(* IEC 61131-3 sources: ICSPrism/benchmarks, 8 files *)

(* ---- harness_test.st ---- *)
FUNCTION_BLOCK Counter
VAR_INPUT
    Increment : INT;
    Reset     : BOOL;
END_VAR
VAR
    Value     : INT;
    TotalCalls: INT;
END_VAR

TotalCalls := TotalCalls + 1;
IF Reset THEN
    Value := 0;
ELSE
    Value := Value + Increment;
END_IF
END_FUNCTION_BLOCK

PROGRAM HarnessTest
VAR_INPUT
    A        : INT;       (* i16 scalar input           *)
    B        : INT;       (* i16 scalar input           *)
    Flag     : BOOL;      (* i8  boolean input          *)
    Index    : INT;       (* i16 used as array index    *)
END_VAR
VAR
    Sum      : INT;       (* A + B each cycle           *)
    Product  : DINT;      (* A * B, wider type          *)
    Buf      : ARRAY[0..15] OF INT;  (* 16-element buffer *)
    C        : Counter;   (* nested function block      *)
    CycleNum : INT;       (* increments every scan      *)
END_VAR

(* Simple deterministic behavior easy to verify *)
CycleNum := CycleNum + 1;
Sum      := A + B;
Product  := A * B;

(* Bounded array write — safe when 0 <= Index <= 15 *)
IF Index >= 0 AND Index <= 15 THEN
    Buf[Index] := Sum;
END_IF

(* Drive the nested counter *)
C(Increment := A, Reset := Flag);

END_PROGRAM

(* ---- harness_test_buggy.st ---- *)
FUNCTION_BLOCK Counter
VAR_INPUT
    Increment : INT;
    Reset     : BOOL;
END_VAR
VAR
    Value     : INT;
    TotalCalls: INT;
END_VAR

TotalCalls := TotalCalls + 1;
IF Reset THEN
    Value := 0;
ELSE
    Value := Value + Increment;
END_IF
END_FUNCTION_BLOCK

PROGRAM HarnessTest
VAR_INPUT
    A        : INT;       (* i16 scalar input           *)
    B        : INT;       (* i16 scalar input           *)
    Flag     : BOOL;      (* i8  boolean input          *)
    Index    : INT;       (* i16 used as array index    *)
END_VAR
VAR
    Sum      : INT;       (* A + B each cycle           *)
    Product  : DINT;      (* A * B, wider type          *)
    Buf      : ARRAY[0..15] OF INT;  (* 16-element buffer *)
    C        : Counter;   (* nested function block      *)
    CycleNum : INT;       (* increments every scan      *)
END_VAR

(* Simple deterministic behavior easy to verify *)
CycleNum := CycleNum + 1;
Sum      := A + B;
Product  := A * B;

(* Bounded array write — safe when 0 <= Index <= 15 *)
IF Index >= 0 OR Index <= 15 THEN
    Buf[Index] := Sum;
END_IF

(* Drive the nested counter *)
C(Increment := A, Reset := Flag);

END_PROGRAM

(* ---- pipeline_controller.st ---- *)
{external}
FUNCTION prism_bug_abort_if : DINT
VAR_INPUT
    should_abort : DINT;
    bug_id       : DINT;
END_VAR
END_FUNCTION

// pipeline_controller — industrial pipeline fill process controller
//
// Bug: Buffer[FillHead] OOB write when FillHead >= 64 (Buffer is [0..63]).
//
// Why this benchmark is decisively harder for input-only fuzzing:
//
//   (1) FillHead is NEVER compared against 64 — it appears only as an array
//       index. trace-cmp has zero visibility into its growth toward 64.
//
//   (2) TWO-DIMENSIONAL ZONE DECAY with 8 zones:
//       FillHead [0,63] is split into 8 zones of 8. Each zone simultaneously
//       requires (PumpRate + ValvePos) AND PipeTemp to be in specific windows.
//       The windows are arranged so that NO fixed (PumpRate, ValvePos, PipeTemp)
//       triple satisfies all 8 zones — and several consecutive zone transitions
//       require coordinated simultaneous changes in multiple inputs.
//
//       Zone 0 [FH  0- 7]: PVsum [60,90]   PipeTemp [50,65]
//       Zone 1 [FH  8-15]: PVsum [80,110]  PipeTemp [62,77]   PVsum up, temp up
//       Zone 2 [FH 16-23]: PVsum [70,100]  PipeTemp [72,87]   PVsum back, temp up
//       Zone 3 [FH 24-31]: PVsum [55, 85]  PipeTemp [65,80]   PVsum down, temp down
//       Zone 4 [FH 32-39]: PVsum [95,125]  PipeTemp [55,70]   PVsum jumps (gap!)
//       Zone 5 [FH 40-47]: PVsum [65, 95]  PipeTemp [78,93]   PVsum down, temp jumps (gap!)
//       Zone 6 [FH 48-55]: PVsum [85,115]  PipeTemp [52,67]   PVsum up, temp folds back (gap!)
//       Zone 7 [FH 56-63]: PVsum [75,105]  PipeTemp [63,78]   PVsum down, temp up
//
//       Critical transitions with NO input overlap between zones:
//         3→4: PVsum must jump from ≤85 to ≥95 (9-unit gap)
//         4→5: PipeTemp must jump from ≤70 to ≥78 while PVsum drops
//         5→6: PipeTemp must drop from ≥78 to ≤67 (fold-back of ~20 units)
//
//   (3) 7 inputs (vs 4 in valve_sequencer) give the custom mutator a richer
//       space: for each zone, PumpRate AND ValvePos AND PipeTemp must be set
//       correctly — three bytes to coordinate, not one.
//
//   (4) Decay is -6 per bad cycle vs +1 advance per 4th qualifying cycle.
//       Random inputs decay FillHead rapidly; only sustained zone-correct
//       inputs allow growth. Without FillHead state signal, the fuzzer cannot
//       know which zone it is in or which transition is approaching.
//
//   (5) Two pre-fill phases (PRIME, FLOW) are guided by trace-cmp and add
//       ~80 cycles of required navigation before FILL begins.
//
// Phase path:
//   IDLE  → Cmd = 1
//   PRIME → PrimeScore >= 8   (every 3rd phase-cycle, combined sum, decay-2) ~30+ cycles
//   FLOW  → FluxScore >= 8    (combined PipeTemp+CoolantRate, halved/11cy)   ~50+ cycles
//   FILL  → FillHead reaches 64 (every 4th qualifying cycle, 8-zone 2D decay) ~300+ cycles
//
// Key variables for state signal: Phase, PrimeScore, FluxScore,
//   FlowAccum, PressAccum, TempAccum, FillHead.
// FillHead is the only one invisible to trace-cmp.
// (PVsum = PumpRate + ValvePos) zone requirements make the state signal
// especially valuable: the fuzzer must know FillHead to know which inputs
// to set, which trace-cmp cannot determine from TempIn comparisons alone.

VAR_GLOBAL CONSTANT
    PHASE_IDLE  : SINT := 0;
    PHASE_PRIME : SINT := 1;
    PHASE_FLOW  : SINT := 2;
    PHASE_FILL  : SINT := 3;
END_VAR

PROGRAM PLC_PRG
VAR_INPUT
    PumpRate    : INT  := 0;
    ValvePos    : INT  := 0;
    PipeTemp    : INT  := 0;
    BackPressure: INT  := 0;
    FeedConc    : INT  := 0;
    CoolantRate : INT  := 0;
    Cmd         : SINT := 0;
END_VAR
VAR
    Ctrl : PipelineCtrl;
END_VAR

Ctrl(
    PumpRate     := PumpRate,
    ValvePos     := ValvePos,
    PipeTemp     := PipeTemp,
    BackPressure := BackPressure,
    FeedConc     := FeedConc,
    CoolantRate  := CoolantRate,
    Cmd          := Cmd
);

END_PROGRAM

FUNCTION_BLOCK PipelineCtrl
VAR_INPUT
    PumpRate    : INT;
    ValvePos    : INT;
    PipeTemp    : INT;
    BackPressure: INT;
    FeedConc    : INT;
    CoolantRate : INT;
    Cmd         : SINT;
END_VAR
VAR_OUTPUT
    Status      : SINT;
END_VAR
VAR
    Phase        : SINT := PHASE_IDLE;
    CycleCount   : INT  := 0;
    // PRIME phase
    PrimeCycles  : INT  := 0;
    PrimeScore   : INT  := 0;
    // FLOW phase
    FluxScore    : INT  := 0;
    FluxSum      : INT  := 0;
    // FILL phase accumulators
    FlowAccum    : INT  := 0;
    PressAccum   : INT  := 0;
    TempAccum    : INT  := 0;
    PhaseCounter : INT  := 0;
    // Hidden OOB counter — NEVER compared against 64, only used as array index
    FillHead     : INT  := 0;
    // OOB write target
    Buffer       : ARRAY[0..63] OF INT;
    PVsum        : INT  := 0;
    i            : INT;
END_VAR

CycleCount := CycleCount + 1;

CASE Phase OF

    PHASE_IDLE:
        IF Cmd = 1 THEN
            FOR i := 0 TO 63 DO
                Buffer[i] := 0;
            END_FOR;
            PrimeCycles  := 0;
            PrimeScore   := 0;
            FluxScore    := 0;
            FlowAccum    := 0;
            PressAccum   := 0;
            TempAccum    := 0;
            PhaseCounter := 0;
            FillHead     := 0;
            PVsum        := 0;
            Phase        := PHASE_PRIME;
        END_IF;

    PHASE_PRIME:
        // Combined PumpRate+BackPressure sum forces simultaneous tuning of
        // two inputs. trace-cmp sees the sum, not individual contributions.
        // Only every 3rd phase-cycle counts; decay-2 forces sustained inputs.
        PrimeCycles := PrimeCycles + 1;
        PVsum := PumpRate + BackPressure;

        IF PrimeCycles MOD 3 = 0 THEN
            IF PVsum >= 80 AND PVsum <= 160 AND ValvePos >= 15 AND ValvePos <= 60 THEN
                PrimeScore := PrimeScore + 1;
            ELSE
                IF PrimeScore > 1 THEN
                    PrimeScore := PrimeScore - 2;
                ELSE
                    PrimeScore := 0;
                END_IF;
            END_IF;
        END_IF;

        IF PrimeScore >= 8 THEN
            Phase := PHASE_FLOW;
        END_IF;

    PHASE_FLOW:
        // Combined PipeTemp + CoolantRate sum partially hides which input is
        // responsible. Halved every 11 global cycles — forces sustained inputs.
        FluxSum := PipeTemp + CoolantRate;

        IF FluxSum >= 80 AND FluxSum <= 160 AND FeedConc >= 20 AND FeedConc <= 70 THEN
            FluxScore := FluxScore + 1;
        ELSE
            IF FluxScore > 1 THEN
                FluxScore := FluxScore - 2;
            ELSE
                FluxScore := 0;
            END_IF;
        END_IF;

        IF CycleCount MOD 11 = 0 AND FluxScore > 0 THEN
            FluxScore := FluxScore / 2;
        END_IF;

        IF FluxScore >= 8 THEN
            Phase := PHASE_FILL;
        END_IF;

    PHASE_FILL:
        PhaseCounter := PhaseCounter + 1;

        // Three accumulator channels — all visible to trace-cmp, which guides
        // the fuzzer into FILL and maintains channel health.

        IF PumpRate >= 40 AND PumpRate <= 90 THEN
            FlowAccum := FlowAccum + 1;
        ELSE
            IF FlowAccum > 1 THEN
                FlowAccum := FlowAccum - 2;
            ELSE
                FlowAccum := 0;
            END_IF;
        END_IF;

        IF BackPressure >= 30 AND BackPressure <= 80 THEN
            PressAccum := PressAccum + 1;
        ELSE
            IF PressAccum > 0 THEN
                PressAccum := PressAccum - 1;
            END_IF;
        END_IF;

        // TempAccum window [50,100] — all zone PipeTemp windows are subsets
        // of this range, so zone requirements always keep TempAccum healthy.
        IF PipeTemp >= 50 AND PipeTemp <= 100 THEN
            TempAccum := TempAccum + 1;
        ELSE
            IF TempAccum > 1 THEN
                TempAccum := TempAccum - 2;
            ELSE
                TempAccum := 0;
            END_IF;
        END_IF;

        // FillHead advances every 4th qualifying cycle.
        // FillHead is NEVER compared against 64 — only appears as array index.
        IF FlowAccum > 6 AND PressAccum > 5 AND TempAccum > 6 THEN
            IF PhaseCounter MOD 4 = 0 THEN
                FillHead := FillHead + 1;
            END_IF;
        END_IF;

        // TWO-DIMENSIONAL ZONE DECAY — the decisive state-signal barrier:
        //
        // FillHead [0,63] is partitioned into 8 zones of 8. Each zone requires
        // BOTH (PumpRate + ValvePos) AND PipeTemp to be in specific windows.
        // These two conditions must be met simultaneously every cycle or FillHead
        // decays by 6 — erasing up to 6 accumulated advances in one bad cycle.
        //
        // Critical transitions (no overlap between adjacent zones):
        //   3→4: PVsum must jump from ≤85 to ≥95 — 9-unit gap, must coordinate
        //         PumpRate AND ValvePos inputs at exactly the right cycle
        //   4→5: PipeTemp must jump ≥8 units while PVsum drops ≥30 units
        //   5→6: PipeTemp must drop ≥11 units (fold-back)
        //
        // trace-cmp instruments PVsum and PipeTemp comparisons but the required
        // windows change with FillHead (state, not input). An input-only fuzzer
        // receives conflicting gradients: e.g., PVsum should be high for zone 4
        // but low for zones 0, 2, 3, 5. Only the key-state signal on FillHead
        // reveals which zone is currently active.
        //
        // A custom mutator with FillHead signal can look up the current zone and
        // set PumpRate, ValvePos, AND PipeTemp precisely — three bytes at once.
        PVsum := PumpRate + ValvePos;

        IF FillHead < 8 THEN
            // Zone 0: PVsum [60,90], PipeTemp [50,65]
            IF PVsum < 60 OR PVsum > 90 OR PipeTemp < 50 OR PipeTemp > 65 THEN
                IF FillHead > 5 THEN
                    FillHead := FillHead - 6;
                ELSE
                    FillHead := 0;
                END_IF;
            END_IF;
        ELSIF FillHead < 16 THEN
            // Zone 1: PVsum [80,110], PipeTemp [62,77]
            IF PVsum < 80 OR PVsum > 110 OR PipeTemp < 62 OR PipeTemp > 77 THEN
                IF FillHead > 5 THEN
                    FillHead := FillHead - 6;
                ELSE
                    FillHead := 0;
                END_IF;
            END_IF;
        ELSIF FillHead < 24 THEN
            // Zone 2: PVsum [70,100], PipeTemp [72,87]
            IF PVsum < 70 OR PVsum > 100 OR PipeTemp < 72 OR PipeTemp > 87 THEN
                IF FillHead > 5 THEN
                    FillHead := FillHead - 6;
                ELSE
                    FillHead := 0;
                END_IF;
            END_IF;
        ELSIF FillHead < 32 THEN
            // Zone 3: PVsum [55,85], PipeTemp [65,80]
            IF PVsum < 55 OR PVsum > 85 OR PipeTemp < 65 OR PipeTemp > 80 THEN
                IF FillHead > 5 THEN
                    FillHead := FillHead - 6;
                ELSE
                    FillHead := 0;
                END_IF;
            END_IF;
        ELSIF FillHead < 40 THEN
            // Zone 4: PVsum [95,125], PipeTemp [55,70]
            // *** GAP from zone 3: PVsum must jump from ≤85 to ≥95 ***
            IF PVsum < 95 OR PVsum > 125 OR PipeTemp < 55 OR PipeTemp > 70 THEN
                IF FillHead > 5 THEN
                    FillHead := FillHead - 6;
                ELSE
                    FillHead := 0;
                END_IF;
            END_IF;
        ELSIF FillHead < 48 THEN
            // Zone 5: PVsum [65,95], PipeTemp [78,93]
            // *** GAP from zone 4: PipeTemp must jump from ≤70 to ≥78 ***
            IF PVsum < 65 OR PVsum > 95 OR PipeTemp < 78 OR PipeTemp > 93 THEN
                IF FillHead > 5 THEN
                    FillHead := FillHead - 6;
                ELSE
                    FillHead := 0;
                END_IF;
            END_IF;
        ELSIF FillHead < 56 THEN
            // Zone 6: PVsum [85,115], PipeTemp [52,67]
            // *** GAP from zone 5: PipeTemp must drop from ≥78 to ≤67 ***
            IF PVsum < 85 OR PVsum > 115 OR PipeTemp < 52 OR PipeTemp > 67 THEN
                IF FillHead > 5 THEN
                    FillHead := FillHead - 6;
                ELSE
                    FillHead := 0;
                END_IF;
            END_IF;
        ELSE
            // Zone 7: PVsum [75,105], PipeTemp [63,78]
            IF PVsum < 75 OR PVsum > 105 OR PipeTemp < 63 OR PipeTemp > 78 THEN
                IF FillHead > 5 THEN
                    FillHead := FillHead - 6;
                ELSE
                    FillHead := 0;
                END_IF;
            END_IF;
        END_IF;

        // OOB write: Buffer is [0..63] (64 elements).
        // FillHead >= 64 writes out of bounds.
        // FillHead appears ONLY here — no comparison against 64 anywhere.
        Buffer[FillHead] := CycleCount;
        IF FillHead > 63 THEN
            prism_bug_abort_if(1, 9001);
        END_IF;

END_CASE;

Status := Phase;

END_FUNCTION_BLOCK

(* ---- pump_controller.st ---- *)
{external}
FUNCTION prism_bug_abort_if : DINT
VAR_INPUT
    should_abort : DINT;
    bug_id       : DINT;
END_VAR
END_FUNCTION

VAR_GLOBAL CONSTANT
    MODE_INIT  : SINT := 0;
    MODE_IDLE  : SINT := 1;
    MODE_ARMED : SINT := 2;
    MODE_RUN   : SINT := 3;
    MODE_FAULT : SINT := 4;
END_VAR

PROGRAM PLC_PRG
VAR_INPUT
    CmdArm    : BOOL := FALSE;
    CmdStart  : BOOL := FALSE;
    CmdReset  : BOOL := FALSE;
    Pressure  : INT := 0;
    Temp      : INT := 0;
END_VAR
VAR
    Controller : PumpController;
END_VAR

Controller(
    CmdArm := CmdArm,
    CmdStart := CmdStart,
    CmdReset := CmdReset,
    Pressure := Pressure,
    Temp := Temp
);

END_PROGRAM

FUNCTION_BLOCK PumpController
VAR_INPUT
    CmdArm    : BOOL;
    CmdStart  : BOOL;
    CmdReset  : BOOL;
    Pressure  : INT;
    Temp      : INT;
END_VAR
VAR
    Mode          : SINT := MODE_INIT;
    CycleCount    : INT := 0;
    PressureScore : INT := 0;
    ArmedCycles   : INT := 0;
    Offset        : INT := 0;
    Buffer        : ARRAY[0..7] OF INT;
    i             : INT;
END_VAR
VAR_OUTPUT
    Status        : SINT;
END_VAR

CycleCount := CycleCount + 1;

CASE Mode OF

    MODE_INIT:
        FOR i := 0 TO 7 DO
            Buffer[i] := 0;
        END_FOR;
        PressureScore := 0;
        ArmedCycles := 0;
        Offset := 0;
        Mode := MODE_IDLE;

    MODE_IDLE:
        IF CmdReset THEN
            PressureScore := 0;
            ArmedCycles := 0;
            Offset := 0;
        END_IF;

        IF CmdArm THEN
            Mode := MODE_ARMED;
            ArmedCycles := 0;
        END_IF;

    MODE_ARMED:
        ArmedCycles := ArmedCycles + 1;

        IF CmdReset THEN
            Mode := MODE_IDLE;
            PressureScore := 0;
            ArmedCycles := 0;
            Offset := 0;
        ELSIF CmdStart AND ArmedCycles >= 3 THEN
            Mode := MODE_RUN;
        END_IF;

    MODE_RUN:
        IF Pressure > 70 THEN
            PressureScore := PressureScore + 1;
        END_IF;

        IF Temp > 50 AND Temp < 60 THEN
            Offset := Offset + 1;
        END_IF;

        IF PressureScore >= 4 THEN
            Buffer[0] := Buffer[0] + 1;
        END_IF;

        IF Buffer[0] > 2 THEN
            Buffer[1] := Buffer[1] + 1;
        END_IF;

        // Deliberate deep bug:
        // Requires entering RUN, then building enough history so Offset becomes large.
        // Input-only fuzzing with frequent resets should struggle more than stateful fuzzing.
        IF Buffer[1] > 1 THEN
            Buffer[Offset] := 1234;
            IF Offset > 7 THEN
                prism_bug_abort_if(1, 9001);
            END_IF;
        END_IF;

        IF CmdReset THEN
            Mode := MODE_IDLE;
            PressureScore := 0;
            ArmedCycles := 0;
            Offset := 0;
        END_IF;

        IF Temp > 90 THEN
            Mode := MODE_FAULT;
        END_IF;

    MODE_FAULT:
        IF CmdReset THEN
            Mode := MODE_IDLE;
            PressureScore := 0;
            ArmedCycles := 0;
            Offset := 0;
        END_IF;

END_CASE;

Status := Mode;

END_FUNCTION_BLOCK

(* ---- scan_cycle_aircraft_oobr.st ---- *)
VAR_GLOBAL CONSTANT
    SS_INITIALIZE: SINT := 0;
    SS_STEP: SINT := 1;
    SS_FIN: SINT := 2;
END_VAR

PROGRAM PLC_PRG
VAR_INPUT
	In: ARRAY[0..7] OF LREAL := [3.0, 2.0, 3.0, 4.0, 1.0, 0.0, -1.0, 2.5];
    ssMethodType: SINT := SS_INITIALIZE;
END_VAR
VAR
	Out: ARRAY[0..1] OF LREAL;
    Code: Code;
END_VAR

// Harness simulation
Code(In, ssMethodType);

END_PROGRAM

FUNCTION_BLOCK Code
VAR_IN_OUT
    InRecv: ARRAY[0..7] OF LREAL;
    ssMethodType: SINT;
END_VAR
VAR
	offset: DWORD;
    CycleCount: INT;
	wGust: LREAL;
    qGust: LREAL;
    iter: INT;
	In: ARRAY[0..64] OF LREAL;
END_VAR
VAR_OUTPUT
    Out: ARRAY[0..1] OF LREAL;
END_VAR

// Complex branching logic
CASE ssMethodType OF

    SS_INITIALIZE:
        // Initialize memory
        FOR iter := 0 TO 64 DO
            In[iter] := 0.0;
        END_FOR;
        ssMethodType := SS_STEP;

    SS_STEP:

        // Copy Inputs
        CycleCount := CycleCount + 1;
        MemCpy(ADR(In), ADR(InRecv), offset);
        wGust := In[0];
        qGust := In[1];

        // Trigger potential memory error (oob read/write)
        // printf('cycle count: %d$N', CycleCount);
        // printf('offset: %d$N', offset);
        IF InRecv[0] > 1.1 AND InRecv[0] < 1.5 AND InRecv[1] > 2 AND InRecv[1] < 2.14 AND InRecv[2] > 5 AND InRecv[2] < 6.5 THEN
            IF CycleCount MOD 2 = 0 THEN
                offset := offset + 10;
            END_IF
        END_IF
        // IF In[CycleCount MOD 64] > 10 THEN
        //     In[CycleCount MOD 64 + 1] := In[CycleCount MOD 64 + 1] * 1.5;
        // ELSE
        //     In[CycleCount MOD 64 + 2] := In[CycleCount MOD 64 + 2] / 0.5;
        // END_IF;

        // More branching
        IF InRecv[2] < 3.5 AND InRecv[2] > 3.01 THEN
            In[3] := In[3] - 0.7;
            IF CycleCount MOD 2 = 0 THEN
                ssMethodType := SS_FIN;
            END_IF
        ELSE
            In[4] := In[4] + 0.8;
            IF In[4] > 1.0 AND IN[4] < 10.0 THEN
                In[5] := In[5] - 0.5;
                // ssMethodType := SS_FIN;
            ELSE
                In[5] := In[5] + 0.5;
                // ssMethodType := SS_INITIALIZE;
            END_IF;
        END_IF;

        // Additional logic for memory error
        IF In[5] < -1.0 THEN
            In[6] := In[6] * 2.0;
            // ssMethodType := SS_FIN;
        ELSE
            In[7] := In[7] / 2.0;
            // offset := offset - 1;
        END_IF;

        // Outputs for Atomic SubSystem: '<Root>/Code 2'
        Out[0] := -0.6385 * wGust;
        Out[1] := (-0.00592 * wGust) + (-0.6571 * qGust);

    SS_FIN:
        // No action
END_CASE;

END_FUNCTION_BLOCK

(* ---- abort_oracle.st ---- *)
{external}
FUNCTION prism_bug_abort_if : DINT
VAR_INPUT
    should_abort : DINT;
    bug_id       : DINT;
END_VAR
END_FUNCTION

PROGRAM abort_oracle
VAR_INPUT
    Trigger : BOOL;
    Value   : INT;
END_VAR
VAR
    Accumulator : DINT;
END_VAR

Accumulator := Accumulator + Value;

IF Trigger THEN
    prism_bug_abort_if(1, 9001);
END_IF;
END_PROGRAM

(* ---- array_lookup.st ---- *)
PROGRAM array_lookup
VAR
    (* Inputs — these are what the fuzzer mutates *)
    index       : INT;      (* array index — dynamic GEP when used to access table *)
    selector    : INT;      (* selects which lookup table to use *)
    bias        : INT;      (* added to the looked-up value *)

    (* Outputs / state *)
    result      : INT;
    safe_result : INT;
    out_a       : INT;
    out_b       : INT;
END_VAR

VAR_TEMP
    table_a     : ARRAY[0..7] OF INT := [10, 20, 30, 40, 50, 60, 70, 80];
    table_b     : ARRAY[0..7] OF INT := [1,  3,  5,  7,  9, 11, 13, 15];
    clamped     : INT;
END_VAR

    (* --- unsafe path: index used directly, dynamic GEP --- *)
    result := table_a[index] + bias;

    (* --- second dynamic GEP on a different table --- *)
    out_a := table_b[index];

    (* --- selector-driven dynamic GEP: two tables, runtime choice --- *)
    IF selector >= 0 AND selector < 8 THEN
        out_b := table_a[selector] + table_b[selector];
    ELSE
        out_b := 0;
    END_IF;

    (* --- safe path: clamped index, should still emit a GEP but
         the analyser may or may not mark it dynamic depending on
         whether it can prove the clamp — useful to compare --- *)
    IF index >= 0 AND index < 8 THEN
        clamped := index;
    ELSE
        clamped := 0;
    END_IF;
    safe_result := table_a[clamped];

END_PROGRAM

(* ---- sanity_test.st ---- *)
PROGRAM sanity_test
VAR_INPUT
    Delta  : INT;
    Reset  : BOOL;
    Enable : BOOL;
END_VAR
VAR
    Accumulator : INT;
    CycleNum    : INT;
    EdgeCount   : INT;
    PrevEnable  : BOOL;
    Armed       : BOOL;
END_VAR

CycleNum := CycleNum + 1;

IF Reset THEN
    Accumulator := 0;
    Armed := FALSE;
ELSE
    IF Enable THEN
        Accumulator := Accumulator + Delta;
    END_IF;

    IF Enable AND NOT PrevEnable THEN
        EdgeCount := EdgeCount + 1;
    END_IF;

    IF Accumulator >= 10 THEN
        Armed := TRUE;
    END_IF;
END_IF;

PrevEnable := Enable;
END_PROGRAM
